# B&R Automation Studio project lab_1_KVBO_07_23_TER
Automation Studio 4.5.2.102

## Configuration Config1

CPU 4PP065.0351-P74, AutomationRuntime D4.52, Build 4.1.2, Vc V4.52.0

### Task classes (Cpu.sw)
```
Cyclic#1:
  Program <- Program.prg
Binaries: udbdef, TCData, ashwd, User, asfw, arconfig, sysconf, Role, ashwac, iomap
Libraries: Library
```

### Hardware
```
4PP065_0351_P74 : 4PP065.0351-P74 v1.0.4.0
  Connector IF5:
    ActivateDevice = 1
  ConfigurationID = labBR
  Simulation = 1
  KeyMappingFile = VC\4PP065_0351_P74.dis
```

- Physical/Config1/4PP065_0351_P74/IoMap.iom: same as Physical/Config1/4PP065_0351_P74/Cpu.per
- Physical/Config1/4PP065_0351_P74/PvMap.vvm: same as Physical/Config1/4PP065_0351_P74/Cpu.per
## Logical view

Binary libraries used (declarations not repeated): operator, runtime, astime, AsIecCon

### Package Logical/Libraries - Global libraries

### Library Logical/Libraries/Library (ANSIC)

#### Library.fun - Exported functions and function blocks
```iecst
{REDUND_ERROR} {REDUND_UNREPLICABLE} FUNCTION_BLOCK FB_Integrator (*TODO: Add your comment here*) (*$GROUP=User,$CAT=User,$GROUPICON=User.png,$CATICON=User.png*)
	VAR_INPUT
		in : {REDUND_UNREPLICABLE} REAL; (*вход интегрирующего звена*)
		out : {REDUND_UNREPLICABLE} REAL; (*выход интегрирующего звена*)
		dt : {REDUND_UNREPLICABLE} REAL; (*шаг расчета (с)*)
	END_VAR
END_FUNCTION_BLOCK

{REDUND_ERROR} {REDUND_UNREPLICABLE} FUNCTION_BLOCK FB_Motor (*TODO: Add your comment here*) (*$GROUP=User,$CAT=User,$GROUPICON=User.png,$CATICON=User.png*)
	VAR_INPUT
		u : {REDUND_UNREPLICABLE} REAL; (*входное напряжение (В)*)
		w : {REDUND_UNREPLICABLE} REAL; (*частота вращения (об\мин)*)
		phi : {REDUND_UNREPLICABLE} REAL; (*положение (рад)*)
		integrator : {REDUND_UNREPLICABLE} FB_Integrator; (*интегратор*)
		Tm : {REDUND_UNREPLICABLE} REAL; (*электромеханическая постоянная времени (с)*)
		ke : {REDUND_UNREPLICABLE} REAL; (*постоянная ЭДС двигателя (В*мин\об)*)
		dt : {REDUND_UNREPLICABLE} REAL; (*шаг расчета (с)*)
	END_VAR
END_FUNCTION_BLOCK

{REDUND_ERROR} {REDUND_UNREPLICABLE} FUNCTION_BLOCK FB_Regulator (*TODO: Add your comment here*) (*$GROUP=User,$CAT=User,$GROUPICON=User.png,$CATICON=User.png*)
	VAR_INPUT
		e : {REDUND_UNREPLICABLE} REAL; (*рассогласование между задающим воздействием и реальной скоростью вращения вала ДПТ (об\мин)*)
		u : {REDUND_UNREPLICABLE} REAL; (*напряжение, подаваемое на вход (В)*)
		k_p : {REDUND_UNREPLICABLE} REAL; (*пропорциональый коэфициент регулятора*)
		k_i : {REDUND_UNREPLICABLE} REAL; (*интегральный коэфициент регулятора*)
		integrator : {REDUND_UNREPLICABLE} FB_Integrator; (*интегратор*)
		iyOld : {REDUND_UNREPLICABLE} REAL; (*хранение предыдущего значения схемы противонакопления*)
		max_abs_value : {REDUND_UNREPLICABLE} REAL; (*граница блока ограничения (В)*)
		dt : {REDUND_UNREPLICABLE} REAL; (*шаг расчета (с)*)
	END_VAR
END_FUNCTION_BLOCK
```

#### FB_Integrator.c
```c
#include <bur/plctypes.h>
#ifdef __cplusplus
	extern "C"
	{
#endif
	#include "Library.h"
#ifdef __cplusplus
	};
#endif
/* TODO: Add your comment here */
void FB_Integrator(struct FB_Integrator* inst)
{
	inst->out += inst->in * inst->dt;
}
```

#### FB_Motor.c
```c
#include <bur/plctypes.h>
#ifdef __cplusplus
	extern "C"
	{
#endif
	#include "Library.h"
#ifdef __cplusplus
	};
#endif
/* TODO: Add your comment here */
void FB_Motor(struct FB_Motor* inst)
{/*
	float delta_w = (inst->u / inst->ke)- inst->w;
	inst->w += delta_w * (inst->dt / inst->Tm);

	inst->integrator.in = inst->w;
	inst->integrator.dt = inst->dt;

	FB_Integrator(&inst->integrator);

	inst->phi = inst->integrator.out;
*/

	inst->integrator.in = (inst->u / inst->ke - inst->w) / inst->Tm;
	inst->integrator.dt = inst->dt;
	FB_Integrator(&inst->integrator);

	inst->w = inst->integrator.out;

	inst->phi = inst->phi + inst->w * 0.10471975512f * inst->dt;
}
```

#### FB_Regulator.c
```c
#include <bur/plctypes.h>
#ifdef __cplusplus
	extern "C"
	{
#endif
	#include "Library.h"
#ifdef __cplusplus
	};
#endif
/* TODO: Add your comment here */

static REAL limit_abs(REAL x, REAL lim)
{
	if (x > lim) return lim;
	if (x < -lim) return -lim;
	return x;

}

void FB_Regulator(struct FB_Regulator* inst)
{/*
	float prop_part = inst->e * inst->k_p;
	if (prop_part > inst->max_abs_value) prop_part = inst->max_abs_value;
	if (prop_part < -inst->max_abs_value) prop_part = -inst->max_abs_value;

	float intteg_input = (inst->e * inst->k_i * inst->dt) + inst->iyOld;
	inst->integrator.in = intteg_input;

	inst->integrator.dt = 1.0f;
	FB_Integrator(&inst->integrator);

	float sum_u = prop_part + inst->integrator.out;

	float limited_u = sum_u;
	if (limited_u > inst->max_abs_value) limited_u = inst->max_abs_value;
	if (limited_u > -inst->max_abs_value) limited_u = -inst->max_abs_value;

	inst->u = limited_u; */

	REAL p_part;
	REAL sum_unlim;

	p_part = limit_abs(inst->k_p*inst->e, inst->max_abs_value);

	inst->integrator.in = inst->k_i * inst->e + inst->iyOld / inst->dt;
	inst->integrator.dt = inst->dt;

	FB_Integrator(&inst->integrator);

	sum_unlim = p_part + inst->integrator.out;

	inst->u = limit_abs(sum_unlim, inst->max_abs_value);

	inst->iyOld = inst->u - sum_unlim;

}
```

### Program Logical/Program (ANSIC)

#### Cyclic.c - Cyclic code
```c
#include <bur/plctypes.h>

#ifdef _DEFAULT_INCLUDES
	#include <AsDefault.h>
#endif

void _CYCLIC ProgramCyclic(void)
{

	counter = counter + fb_motor.dt;
	if (counter  >= 60.0f) counter = 0.0f;
	if (counter > 20.0f && counter < 40.0f) Speed = 60.0f;
	else {
		Speed = 0.0f;
	}
	fb_controller.e = Speed - fb_motor.w;

	FB_Regulator(&fb_controller);

	fb_motor.u = fb_controller.u;
	fb_motor2.u = Speed*fb_motor2.ke;

	FB_Motor(&fb_motor2);
	FB_Motor(&fb_motor);
}
```

#### Init.c - Initialization code
```c
#include <bur/plctypes.h>

#ifdef _DEFAULT_INCLUDES
	#include <AsDefault.h>
#endif

void _INIT ProgramInit(void)
{
	float dt = 0.01f;
	float Tj = 0.3f;

	fb_controller.max_abs_value = 24.0f;
	fb_controller.dt = dt;
	fb_controller.iyOld = 0.0f;
	fb_controller.integrator.out = 0.0f;

	fb_motor.ke = 0.01f;
	fb_motor.Tm = 0.05f;
	fb_motor.dt = dt;
	fb_motor.w = 0.0f;
	fb_motor.phi = 0.0f;
	fb_motor.integrator.out = 0.0f;

	fb_motor2.ke = 0.01f;
	fb_motor2.Tm = 0.05f;
	fb_motor2.dt = dt;
	fb_motor2.w = 0.0f;
	fb_motor2.phi = 0.0f;
	fb_motor2.integrator.out = 0.0f;

	fb_controller.k_p = fb_motor.ke * fb_motor.Tm / Tj;
	fb_controller.k_i = fb_motor.ke / Tj;

	counter = 0.0f;
	Speed = 0.0f;
	Enable = 1;
}
```

#### Exit.c - Exit code
```c
#include <bur/plctypes.h>

#ifdef _DEFAULT_INCLUDES
	#include <AsDefault.h>
#endif

void _EXIT ProgramExit(void)
{

}
```

#### Variables.var - Local variables
```iecst
VAR
	fb_controller : FB_Regulator;
	fb_motor : FB_Motor;
	Speed : REAL;
	Enable : BOOL;
	counter : REAL;
	fb_motor2 : FB_Motor;
END_VAR
```
